(* IEC 61131-3 sources: rusty/tests/lit/cfc/blocks/function_void, 2 files *)

(* ---- main.st ---- *)
FUNCTION main : DINT
    function_void();
    // CHECK: result = 6
    printf('result = %d$N', function_void.localOut);
END_FUNCTION

(* ---- myVoid.st ---- *)
FUNCTION myVoid
VAR_INPUT
    in : DINT;
END_VAR
VAR_OUTPUT
    out : DINT;
END_VAR
    out := in * 2;
END_FUNCTION
